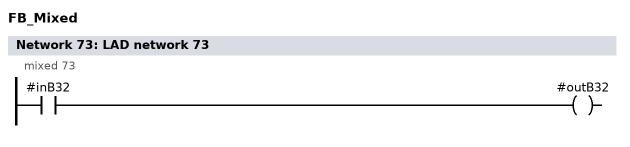
   RUNG wire#powerrail
      Contact( #inB32 )
      Coil( #outB32 )
   END_RUNG
   // the same network as SCL:
   #outB32 := #inB32;
END_REGION

REGION Network 74 (FBD): FBD network 74
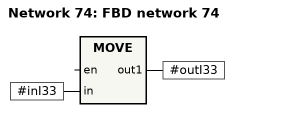
   #outI33 := #inI33;
END_REGION

REGION Network 75 (SCL): SCL network 75
   #tI74 := #inI34 + #cI14;
           IF #inB34 THEN
               #outR14 := #inR14 * 2.0;
           END_IF;
END_REGION

REGION Network 76: LAD network 76
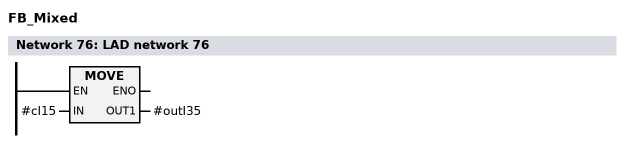
   RUNG wire#powerrail
      Move(in := #cI15, out1 => #outI35)
   END_RUNG
   // the same network as SCL:
   #outI35 := #cI15;
END_REGION

REGION Network 77 (FBD): FBD network 77
   // mixed 77
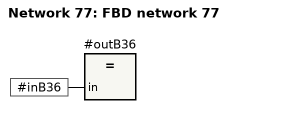
   #outB36 := #inB36;
END_REGION

REGION Network 78 (SCL): SCL network 78
   #tI77 := #inI37 + #cI17;
           IF #inB37 THEN
               #outR17 := #inR17 * 2.0;
           END_IF;
END_REGION

REGION Network 79: LAD network 79
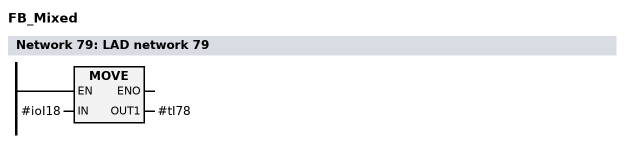
   RUNG wire#powerrail
      Move(in := #ioI18, out1 => #tI78)
   END_RUNG
   // the same network as SCL:
   #tI78 := #ioI18;
END_REGION

REGION Network 80 (FBD): FBD network 80
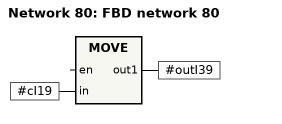
   #outI39 := #cI19;
END_REGION

REGION Network 81 (SCL): SCL network 81
   // mixed 81
   #tI80 := #inI0 + #cI20;
           IF #inB0 THEN
               #outR0 := #inR0 * 2.0;
           END_IF;
END_REGION

REGION Network 82: LAD network 82
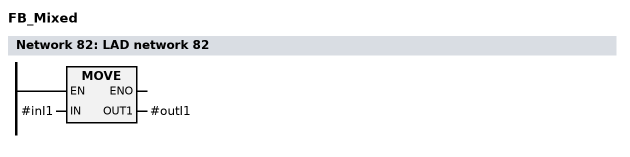
   RUNG wire#powerrail
      Move(in := #inI1, out1 => #outI1)
   END_RUNG
   // the same network as SCL:
   #outI1 := #inI1;
END_REGION

REGION Network 83 (FBD): FBD network 83
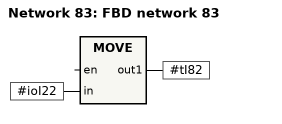
   #tI82 := #ioI22;
END_REGION

REGION Network 84 (SCL): SCL network 84
   #tI83 := #inI3 + #cI23;
           IF #inB3 THEN
               #outR3 := #inR3 * 2.0;
           END_IF;
END_REGION

REGION Network 85: LAD network 85
   // mixed 85
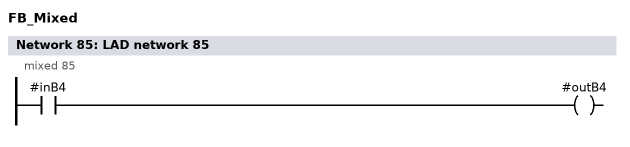
   RUNG wire#powerrail
      Contact( #inB4 )
      Coil( #outB4 )
   END_RUNG
   // the same network as SCL:
   #outB4 := #inB4;
END_REGION

REGION Network 86 (FBD): FBD network 86
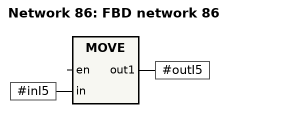
   #outI5 := #inI5;
END_REGION

REGION Network 87 (SCL): SCL network 87
   #tI86 := #inI6 + #cI26;
           IF #inB6 THEN
               #outR6 := #inR6 * 2.0;
           END_IF;
END_REGION

REGION Network 88: LAD network 88
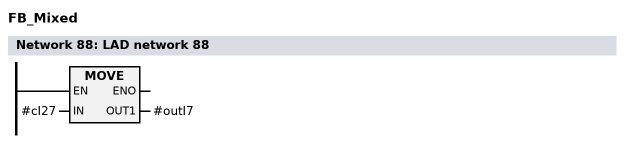
   RUNG wire#powerrail
      Move(in := #cI27, out1 => #outI7)
   END_RUNG
   // the same network as SCL:
   #outI7 := #cI27;
END_REGION

REGION Network 89 (FBD): FBD network 89
   // mixed 89
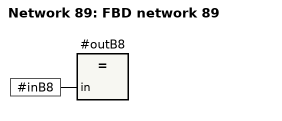
   #outB8 := #inB8;
END_REGION

REGION Network 90 (SCL): SCL network 90
   #tI89 := #inI9 + #cI29;
           IF #inB9 THEN
               #outR9 := #inR9 * 2.0;
           END_IF;
END_REGION

REGION Network 91: LAD network 91
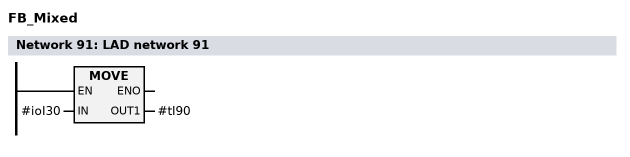
   RUNG wire#powerrail
      Move(in := #ioI30, out1 => #tI90)
   END_RUNG
   // the same network as SCL:
   #tI90 := #ioI30;
END_REGION

REGION Network 92 (FBD): FBD network 92
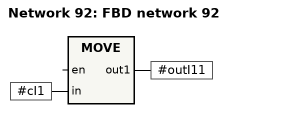
   #outI11 := #cI1;
END_REGION

REGION Network 93 (SCL): SCL network 93
   // mixed 93
   #tI92 := #inI12 + #cI2;
           IF #inB12 THEN
               #outR12 := #inR12 * 2.0;
           END_IF;
END_REGION

REGION Network 94: LAD network 94
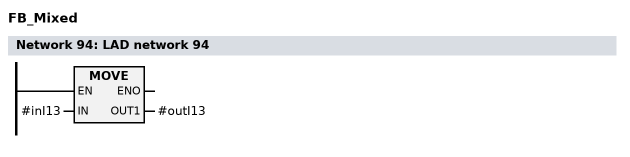
   RUNG wire#powerrail
      Move(in := #inI13, out1 => #outI13)
   END_RUNG
   // the same network as SCL:
   #outI13 := #inI13;
END_REGION

REGION Network 95 (FBD): FBD network 95
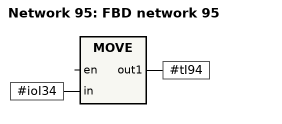
   #tI94 := #ioI34;
END_REGION

REGION Network 96 (SCL): SCL network 96
   #tI95 := #inI15 + #cI5;
           IF #inB15 THEN
               #outR15 := #inR15 * 2.0;
           END_IF;
END_REGION

REGION Network 97: LAD network 97
   // mixed 97
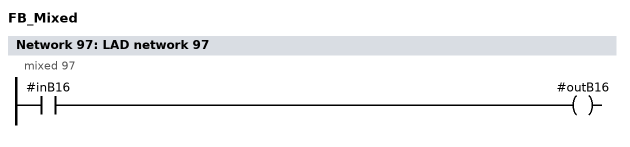
   RUNG wire#powerrail
      Contact( #inB16 )
      Coil( #outB16 )
   END_RUNG
   // the same network as SCL:
   #outB16 := #inB16;
END_REGION

REGION Network 98 (FBD): FBD network 98
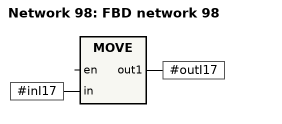
   #outI17 := #inI17;
END_REGION

REGION Network 99 (SCL): SCL network 99
   #tI98 := #inI18 + #cI8;
           IF #inB18 THEN
               #outR18 := #inR18 * 2.0;
           END_IF;
END_REGION

REGION Network 100: LAD network 100
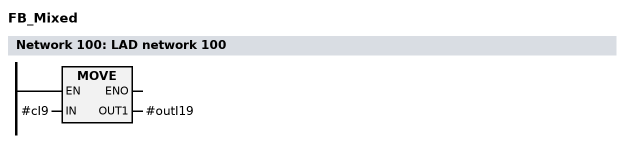
   RUNG wire#powerrail
      Move(in := #cI9, out1 => #outI19)
   END_RUNG
   // the same network as SCL:
   #outI19 := #cI9;
END_REGION

REGION Network 101 (FBD): FBD network 101
   // mixed 101
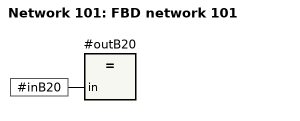
   #outB20 := #inB20;
END_REGION

REGION Network 102 (SCL): SCL network 102
   #tI1 := #inI21 + #cI11;
           IF #inB21 THEN
               #outR1 := #inR1 * 2.0;
           END_IF;
END_REGION

REGION Network 103: LAD network 103
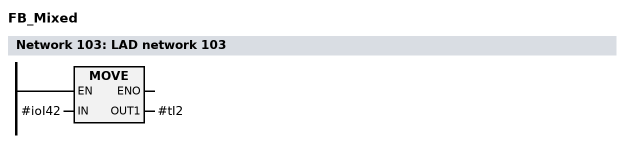
   RUNG wire#powerrail
      Move(in := #ioI42, out1 => #tI2)
   END_RUNG
   // the same network as SCL:
   #tI2 := #ioI42;
END_REGION

REGION Network 104 (FBD): FBD network 104
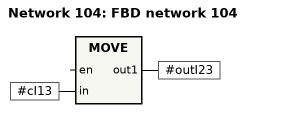
   #outI23 := #cI13;
END_REGION

REGION Network 105 (SCL): SCL network 105
   // mixed 105
   #tI4 := #inI24 + #cI14;
           IF #inB24 THEN
               #outR4 := #inR4 * 2.0;
           END_IF;
END_REGION

REGION Network 106: LAD network 106
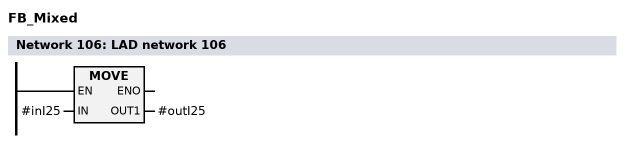
   RUNG wire#powerrail
      Move(in := #inI25, out1 => #outI25)
   END_RUNG
   // the same network as SCL:
   #outI25 := #inI25;
END_REGION

REGION Network 107 (FBD): FBD network 107
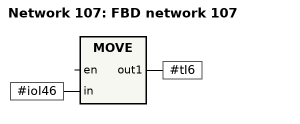
   #tI6 := #ioI46;
END_REGION

REGION Network 108 (SCL): SCL network 108
   #tI7 := #inI27 + #cI17;
           IF #inB27 THEN
               #outR7 := #inR7 * 2.0;
           END_IF;
END_REGION

REGION Network 109: LAD network 109
   // mixed 109
